FUNCTION_BLOCK FB_AnalogInput (* Migrated from IEC 61131-3 ST *)
  (* Standard: 61499-2 *)
  (* Version 1.0, 2026-11-06, st2fb *)
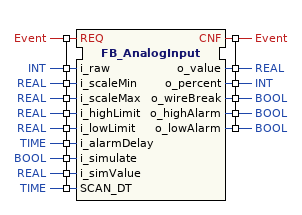
  EVENT_INPUT
    REQ WITH i_raw, i_scaleMin, i_scaleMax, i_highLimit, i_lowLimit, i_alarmDelay, i_simulate, i_simValue, SCAN_DT;
  END_EVENT
  EVENT_OUTPUT
    CNF WITH o_value, o_percent, o_wireBreak, o_highAlarm, o_lowAlarm;
  END_EVENT
  VAR_INPUT
    i_raw : INT;
    i_scaleMin : REAL;
    i_scaleMax : REAL;
    i_highLimit : REAL;
    i_lowLimit : REAL;
    i_alarmDelay : TIME;
    i_simulate : BOOL;
    i_simValue : REAL;
    SCAN_DT : TIME;
  END_VAR
  VAR_OUTPUT
    o_value : REAL;
    o_percent : INT;
    o_wireBreak : BOOL;
    o_highAlarm : BOOL;
    o_lowAlarm : BOOL;
  END_VAR
  VAR
    ST2FB_NOW : TIME := T#0s;
    statLastGood : REAL := 0.0;
    statDelay : TIME := T#0s;
    statTiming : BOOL := FALSE;
    tempNorm : REAL := 0.0;
    tempScaled : REAL := 0.0;
    tempBreak : BOOL := FALSE;
    tempHigh : BOOL := FALSE;
    tempLow : BOOL := FALSE;
    H_IN : BOOL := FALSE;
    H_PT : TIME := T#0s;
    H_Q : BOOL := FALSE;
    H_ET : TIME := T#0s;
    H_STATE : INT := 0;
    H_PREV_IN : BOOL := FALSE;
    H_START_TIME : TIME := T#0s;
    L_IN : BOOL := FALSE;
    L_PT : TIME := T#0s;
    L_Q : BOOL := FALSE;
    L_ET : TIME := T#0s;
    L_STATE : INT := 0;
    L_PREV_IN : BOOL := FALSE;
    L_START_TIME : TIME := T#0s;
    B_IN : BOOL := FALSE;
    B_PT : TIME := T#0s;
    B_Q : BOOL := FALSE;
    B_ET : TIME := T#0s;
    B_STATE : INT := 0;
    B_PREV_IN : BOOL := FALSE;
    B_START_TIME : TIME := T#0s;
  END_VAR
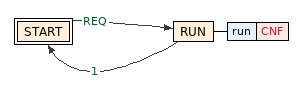
  EC_STATES
    START;
    RUN : run -> CNF;
  END_STATES
  EC_TRANSITIONS
    START TO RUN := REQ;
    RUN TO START := 1;
  END_TRANSITIONS
  ALGORITHM run IN ST:
ST2FB_NOW := ST2FB_NOW + SCAN_DT;
tempNorm := (INT_TO_REAL(i_raw) - 0.0) / (27648.0 - 0.0);
tempScaled := tempNorm * (i_scaleMax - i_scaleMin) + i_scaleMin;

IF NOT statTiming THEN
  statDelay := i_alarmDelay;
END_IF;

tempBreak := i_raw = 32767;
B_IN := tempBreak;
B_PT := statDelay;
IF (B_STATE = 0) AND NOT B_PREV_IN AND B_IN THEN
  B_STATE := 1;
  B_Q := FALSE;
  B_START_TIME := ST2FB_NOW;
ELSE
  IF NOT B_IN THEN
    B_ET := T#0s;
    B_Q := FALSE;
    B_STATE := 0;
  ELSIF B_STATE = 1 THEN
    IF B_START_TIME + B_PT <= ST2FB_NOW THEN
      B_STATE := 2;
      B_Q := TRUE;
      B_ET := B_PT;
    ELSE
      B_ET := ST2FB_NOW - B_START_TIME;
    END_IF;
  END_IF;
END_IF;
B_PREV_IN := B_IN;
o_wireBreak := B_Q;
IF i_raw <> 32767 THEN
  statLastGood := tempScaled;
END_IF;

IF i_simulate THEN
  o_value := i_simValue;
ELSE
  o_value := statLastGood;
END_IF;
o_percent := REAL_TO_INT(100.0 * LIMIT(0.0, tempNorm, 1.0));

tempHigh := o_value > i_highLimit;
tempLow := o_value < i_lowLimit;

H_IN := tempHigh;
H_PT := statDelay;
IF (H_STATE = 0) AND NOT H_PREV_IN AND H_IN THEN
  H_STATE := 1;
  H_Q := FALSE;
  H_START_TIME := ST2FB_NOW;
ELSE
  IF NOT H_IN THEN
    H_ET := T#0s;
    H_Q := FALSE;
    H_STATE := 0;
  ELSIF H_STATE = 1 THEN
    IF H_START_TIME + H_PT <= ST2FB_NOW THEN
      H_STATE := 2;
      H_Q := TRUE;
      H_ET := H_PT;
    ELSE
      H_ET := ST2FB_NOW - H_START_TIME;
    END_IF;
  END_IF;
END_IF;
H_PREV_IN := H_IN;
o_highAlarm := H_Q;

L_IN := tempLow;
L_PT := statDelay;
IF (L_STATE = 0) AND NOT L_PREV_IN AND L_IN THEN
  L_STATE := 1;
  L_Q := FALSE;
  L_START_TIME := ST2FB_NOW;
ELSE
  IF NOT L_IN THEN
    L_ET := T#0s;
    L_Q := FALSE;
    L_STATE := 0;
  ELSIF L_STATE = 1 THEN
    IF L_START_TIME + L_PT <= ST2FB_NOW THEN
      L_STATE := 2;
      L_Q := TRUE;
      L_ET := L_PT;
    ELSE
      L_ET := ST2FB_NOW - L_START_TIME;
    END_IF;
  END_IF;
END_IF;
L_PREV_IN := L_IN;
o_lowAlarm := L_Q;

statTiming := tempBreak OR tempHigh OR tempLow;
  END_ALGORITHM
END_FUNCTION_BLOCK
